(* IEC 61131-3 sources: Caravan/Archiv/12-04-19/Stations/Terminal/HMI/Network/STDCommunicationToPLC, 1 file *)

(* ---- ONE_STDCommunicationToPLC_Table.st ---- *)
#define OBJECTS_CONFIG

#include "..\..\Class\_AlarmX0Para\_AlarmX0Para.h"
#include "..\..\Class\DataManager\DataManager.h"
//Define part of class DataManagerFIFO
#define MEMORY_Mark_DataMngFiFo    8
#include "..\..\Class\TCPCommunication\TCPCommunication.h"
#include "..\..\Class\TCPCommunication\SalamanderDelay.h"
#include "..\..\Class\TCPCommunicationLogViewer\TCPCommunicationLogViewer.h"

FUNCTION GLOBAL TAB ONE_STDCommunicationToPLC
-1$UINT, 0$UINT,
1$UINT, 0$UINT,

18$UDINT,
TO_UDINT(800276940), "_AlarmX0Para", 0$UINT, 11$UINT, 1$UINT,
TO_UDINT(3900434542), "_CheckOnlineStatus", 1$UINT, 3$UINT, 1$UINT,
TO_UDINT(916194998), "_CheckSum", 1$UINT, 0$UINT, 1$UINT,
TO_UDINT(2980745877), "_MyIO", 0$UINT, 3$UINT, 0$UINT,
TO_UDINT(3043040051), "_ScrollArea", 0$UINT, 15$UINT, 0$UINT,
TO_UDINT(2779823616), "_ScrollArea2", 0$UINT, 8$UINT, 0$UINT,
TO_UDINT(794617671), "CriticalSection", 0$UINT, 4$UINT, 10$UINT,
TO_UDINT(4008337867), "DataManager", 1$UINT, 0$UINT, 1$UINT,
TO_UDINT(2873804345), "DataManagerFIFO", 1$UINT, 0$UINT, 10$UINT,
TO_UDINT(2393054465), "DataManagerPriority", 1$UINT, 0$UINT, 1$UINT,
TO_UDINT(2602835227), "GetTaskHandle", 0$UINT, 2$UINT, 1$UINT,
TO_UDINT(2225119864), "MerkerEx", 1$UINT, 21$UINT, 2$UINT,
TO_UDINT(3534980377), "RamRingBuffer", 1$UINT, 1$UINT, 1$UINT,
TO_UDINT(1850111279), "String", 1$UINT, 10$UINT, 1$UINT,
TO_UDINT(2898603620), "StringInternal", 1$UINT, 82$UINT, 0$UINT,
TO_UDINT(3704218787), "TCPCommunication", 1$UINT, 14$UINT, 1$UINT,
TO_UDINT(185738949), "TCPCommunicationLogViewer", 1$UINT, 4$UINT, 1$UINT,
TO_UDINT(3232495061), "VirtualBaseInit", 1$UINT, 3$UINT, 0$UINT,

_NO_ATTR, TO_UDINT(2307429966), "ALARMCOMMUNICATION_HMI",

_NO_ATTR, TO_UDINT(4100950075), "CHECKCOMM",

1$UINT, TO_UDINT(1793796099), "STDTCPCOMMUNICATIONTOMC1\CHECKSUM",

1$UINT, TO_UDINT(494624950), "STDDATAMANAGERTOMC1\DATAMANAGERPRIORITY\DATAMANAGERFIFO_PRIO0\SECTION",
1$UINT, TO_UDINT(167802101), "STDDATAMANAGERTOMC1\DATAMANAGERPRIORITY\DATAMANAGERFIFO_PRIO1\SECTION",
1$UINT, TO_UDINT(864897072), "STDDATAMANAGERTOMC1\DATAMANAGERPRIORITY\DATAMANAGERFIFO_PRIO2\SECTION",
1$UINT, TO_UDINT(620125299), "STDDATAMANAGERTOMC1\DATAMANAGERPRIORITY\DATAMANAGERFIFO_PRIO3\SECTION",
1$UINT, TO_UDINT(1083650490), "STDDATAMANAGERTOMC1\DATAMANAGERPRIORITY\DATAMANAGERFIFO_PRIO4\SECTION",
1$UINT, TO_UDINT(1475094009), "STDDATAMANAGERTOMC1\DATAMANAGERPRIORITY\DATAMANAGERFIFO_PRIO5\SECTION",
1$UINT, TO_UDINT(1851857212), "STDDATAMANAGERTOMC1\DATAMANAGERPRIORITY\DATAMANAGERFIFO_PRIO6\SECTION",
1$UINT, TO_UDINT(2031750527), "STDDATAMANAGERTOMC1\DATAMANAGERPRIORITY\DATAMANAGERFIFO_PRIO7\SECTION",
1$UINT, TO_UDINT(2795750062), "STDDATAMANAGERTOMC1\DATAMANAGERPRIORITY\DATAMANAGERFIFO_PRIO8\SECTION",
1$UINT, TO_UDINT(2983778029), "STDDATAMANAGERTOMC1\DATAMANAGERPRIORITY\DATAMANAGERFIFO_PRIO9\SECTION",

_NO_ATTR, TO_UDINT(968784990), "STDDATAMANAGERTOMC1",

1$UINT, TO_UDINT(1138546362), "STDDATAMANAGERTOMC1\DATAMANAGERPRIORITY\DATAMANAGERFIFO_PRIO0",
1$UINT, TO_UDINT(886826540), "STDDATAMANAGERTOMC1\DATAMANAGERPRIORITY\DATAMANAGERFIFO_PRIO1",
1$UINT, TO_UDINT(2916267926), "STDDATAMANAGERTOMC1\DATAMANAGERPRIORITY\DATAMANAGERFIFO_PRIO2",
1$UINT, TO_UDINT(3671426816), "STDDATAMANAGERTOMC1\DATAMANAGERPRIORITY\DATAMANAGERFIFO_PRIO3",
1$UINT, TO_UDINT(1152455331), "STDDATAMANAGERTOMC1\DATAMANAGERPRIORITY\DATAMANAGERFIFO_PRIO4",
1$UINT, TO_UDINT(867574325), "STDDATAMANAGERTOMC1\DATAMANAGERPRIORITY\DATAMANAGERFIFO_PRIO5",
1$UINT, TO_UDINT(2864673679), "STDDATAMANAGERTOMC1\DATAMANAGERPRIORITY\DATAMANAGERFIFO_PRIO6",
1$UINT, TO_UDINT(3719840537), "STDDATAMANAGERTOMC1\DATAMANAGERPRIORITY\DATAMANAGERFIFO_PRIO7",
1$UINT, TO_UDINT(1292328584), "STDDATAMANAGERTOMC1\DATAMANAGERPRIORITY\DATAMANAGERFIFO_PRIO8",
1$UINT, TO_UDINT(973106718), "STDDATAMANAGERTOMC1\DATAMANAGERPRIORITY\DATAMANAGERFIFO_PRIO9",

1$UINT, TO_UDINT(2505094980), "STDDATAMANAGERTOMC1\DATAMANAGERPRIORITY",

1$UINT, TO_UDINT(1712597188), "STDDATAMANAGERTOMC1\DATAMNGGETTASKHANDLE1",

1$UINT, TO_UDINT(2307201355), "STDTCPCOMMUNICATIONTOMC1\RAMRINGMERKEREX",
1$UINT, TO_UDINT(569575462), "STDTCPCOMMUNICATIONTOMC1\THREADNAME\MERKEREX0",

1$UINT, TO_UDINT(2727999187), "STDTCPCOMMUNICATIONTOMC1\RAMRINGBUFFER",

1$UINT, TO_UDINT(832950765), "STDTCPCOMMUNICATIONTOMC1\THREADNAME",

_NO_ATTR, TO_UDINT(2516610500), "STDTCPCOMMUNICATIONTOMC1",

_NO_ATTR, TO_UDINT(705022640), "STDTCPCOMMUNICATIONLOGVIEWER1",

//Internal connections
0$UDINT,
27$UDINT,
TO_UDINT(13), "DataMngGetTaskHandle1", TO_UDINT(25),
TO_UDINT(13), "DataManagerPriority", TO_UDINT(24),
TO_UDINT(14), "Section", TO_UDINT(3),
TO_UDINT(15), "Section", TO_UDINT(4),
TO_UDINT(16), "Section", TO_UDINT(5),
TO_UDINT(17), "Section", TO_UDINT(6),
TO_UDINT(18), "Section", TO_UDINT(7),
TO_UDINT(19), "Section", TO_UDINT(8),
TO_UDINT(20), "Section", TO_UDINT(9),
TO_UDINT(21), "Section", TO_UDINT(10),
TO_UDINT(22), "Section", TO_UDINT(11),
TO_UDINT(23), "Section", TO_UDINT(12),
TO_UDINT(24), "DataManagerFiFo_Prio0", TO_UDINT(14),
TO_UDINT(24), "DataManagerFiFo_Prio1", TO_UDINT(15),
TO_UDINT(24), "DataManagerFiFo_Prio2", TO_UDINT(16),
TO_UDINT(24), "DataManagerFiFo_Prio3", TO_UDINT(17),
TO_UDINT(24), "DataManagerFiFo_Prio4", TO_UDINT(18),
TO_UDINT(24), "DataManagerFiFo_Prio5", TO_UDINT(19),
TO_UDINT(24), "DataManagerFiFo_Prio6", TO_UDINT(20),
TO_UDINT(24), "DataManagerFiFo_Prio7", TO_UDINT(21),
TO_UDINT(24), "DataManagerFiFo_Prio8", TO_UDINT(22),
TO_UDINT(24), "DataManagerFiFo_Prio9", TO_UDINT(23),
TO_UDINT(29), "MerkerEx0", TO_UDINT(27),
TO_UDINT(30), "RamRingBuffer", TO_UDINT(28),
TO_UDINT(30), "RamRingMerkerEx", TO_UDINT(26),
TO_UDINT(30), "CheckSum", TO_UDINT(2),
TO_UDINT(30), "ThreadName", TO_UDINT(29),
0$UDINT,
7$UDINT,
TO_UDINT(1), "toTCPComm", TO_UDINT(30), "ClassSvr",
TO_UDINT(1), "AlarmCommunication", TO_UDINT(0), "ClassSvr",
TO_UDINT(13), "coTCPCommunication", TO_UDINT(30), "ClassSvr",
TO_UDINT(28), "Data", TO_UDINT(26), "m_udLength",
TO_UDINT(29), "DataBuffer", TO_UDINT(27), "m_udLength",
TO_UDINT(30), "coDataMng", TO_UDINT(13), "ClassSvr",
TO_UDINT(31), "coTCPCommunication", TO_UDINT(30), "ClassSvr",

//Initialization values
0$UDINT,
13$UDINT,
TO_UDINT(0), "Config", TO_UDINT(10000),//|STDCommunicationToPLC.AlarmCommunication_HMI.Config;
TO_UDINT(1), "DelayTime", TO_UDINT(20000),//|STDCommunicationToPLC.CheckComm.DelayTime;
TO_UDINT(13), "AcceptOfflineJobs", TO_UDINT(1),//|STDCommunicationToPLC.STDDataManagerToMC1.AcceptOfflineJobs;
TO_UDINT(26), "ThreadSafe", TO_UDINT(0),//|STDCommunicationToPLC.STDTCPCommunicationToMC1\RamRingMerkerEx.ThreadSafe;
TO_UDINT(27), "ThreadSafe", TO_UDINT(0),//|STDCommunicationToPLC.ThreadName\STDTCPCommunicationToMC1\MerkerEx0.ThreadSafe;
TO_UDINT(29), "SingleRealloc", TO_UDINT(1),//|STDCommunicationToPLC.STDTCPCommunicationToMC1\ThreadName.SingleRealloc;
TO_UDINT(30), "ComPort", TO_UDINT(500),//|STDCommunicationToPLC.STDTCPCommunicationToMC1.ComPort;
TO_UDINT(30), "LogEnable", TO_UDINT(0),//|STDCommunicationToPLC.STDTCPCommunicationToMC1.LogEnable;
TO_UDINT(30), "DeactivateCom", TO_UDINT(0),//|STDCommunicationToPLC.STDTCPCommunicationToMC1.DeactivateCom;
TO_UDINT(30), "SizeOfComBuffers", TO_UDINT(2MB),//|STDCommunicationToPLC.STDTCPCommunicationToMC1.SizeOfComBuffers;
TO_UDINT(31), "VerticalLevel", TO_UDINT(1),//|STDCommunicationToPLC.STDTCPCommunicationLogViewer1.VerticalLevel;
TO_UDINT(31), "LineWidth", TO_UDINT(0),//|STDCommunicationToPLC.STDTCPCommunicationLogViewer1.LineWidth;
TO_UDINT(31), "ExtendedScrollBar", TO_UDINT(0),//|STDCommunicationToPLC.STDTCPCommunicationLogViewer1.ExtendedScrollBar;

//Symbolic initialization values
0$UDINT,
0$UDINT,

//Initialization of string values
0$UDINT,
0$UDINT,

//Configuration of tasks (RealTime, Cyclic, Background)
0$UDINT,
1$UDINT,
TO_UDINT(25), (1000)$UDINT, 4194303$DINT, 	//STDDATAMANAGERTOMC1\DATAMNGGETTASKHANDLE1

0$UDINT,
4$UDINT,
TO_UDINT(1), (50)$UDINT, 4194303$DINT, 	//CHECKCOMM
TO_UDINT(25), (1000)$UDINT, 4194303$DINT, 	//STDDATAMANAGERTOMC1\DATAMNGGETTASKHANDLE1
TO_UDINT(30), (100)$UDINT, 4194303$DINT, 	//STDTCPCOMMUNICATIONTOMC1
TO_UDINT(31), (1)$UDINT, 4194303$DINT, 	//STDTCPCOMMUNICATIONLOGVIEWER1

0$UDINT,
1$UDINT,
TO_UDINT(25), (1000)$UDINT, 4194303$DINT, 	//STDDATAMANAGERTOMC1\DATAMNGGETTASKHANDLE1

//External connections
0$UDINT,
4$UDINT,
TO_UDINT(30), "coStationToConnect", C_TRY, TO_UDINT(2925151108), "GlobalScreen1","IP4Communication",
TO_UDINT(31), "Lse", C_DIR, TO_UDINT(299963966), "Lse","Lse",
TO_UDINT(31), "SysDate", C_DIR, TO_UDINT(3035062039), "SysDateTime","SysDate",
TO_UDINT(31), "SysTime", C_DIR, TO_UDINT(3035062039), "SysDateTime","SysTime",

//Magic internal connections
0$UDINT,
0$UDINT,

//Configuration of timeslots of tasks (RealTime, Cyclic)
#ifdef __LSLLDR_TIMESLOTS__
0$UDINT,
0$UDINT,

0$UDINT,
0$UDINT,

#endif //__LSLLDR_TIMESLOTS__

//MultiMaster connections
#ifdef __LSLLDR_MULTIMASTER__
0$UDINT,
0$UDINT,
#endif //__LSLLDR_MULTIMASTER__

//Configuration for task ID (RealTime, CyclicTime)
#ifdef __LSLLDR_TASKID__
"\\\\TASKS2  "
0$UDINT,
1$UDINT,
(0)$UDINT, 	//STDDATAMANAGERTOMC1\DATAMNGGETTASKHANDLE1

0$UDINT,
4$UDINT,
(0)$UDINT, 	//CHECKCOMM
(0)$UDINT, 	//STDDATAMANAGERTOMC1\DATAMNGGETTASKHANDLE1
(0)$UDINT, 	//STDTCPCOMMUNICATIONTOMC1
(0)$UDINT, 	//STDTCPCOMMUNICATIONLOGVIEWER1

0$UDINT,
1$UDINT,
(0)$UDINT, 	//STDDATAMANAGERTOMC1\DATAMNGGETTASKHANDLE1

#endif //__LSLLDR_TASKID__

END_FUNCTION
